// TIA Portal V21 export
// export: Created 2026-11-09T01:07:26.0249752Z, ExportSetting WithDefaults, DisplayName Totally Integrated Automation Portal, DisplayVersion V21 Update 3, DisplayName STEP 7 Professional, DisplayVersion V21 Update 3, DisplayName STEP 7 Safety, DisplayVersion V21, DisplayName Tech WebApplication, DisplayVersion V21, DisplayName WinCC Basic/Comfort/Advanced, DisplayVersion V21 Update 3, DisplayName WinCC Unified, DisplayVersion V21 Update 3
FUNCTION_BLOCK "FB_Motor"   // FB2, SCL
{ S7_Optimized_Access := 'TRUE' }
// stored: AutoNumber true, IsIECCheckEnabled false, IsRetainMemResEnabled false, MemoryReserve 100, SetENOAutomatically false, UDAEnableTagReadback false
   VAR_INPUT
      motor : "UDT_Motor";
   END_VAR
   VAR_OUTPUT
      running : Bool;
   END_VAR
BEGIN
   #running := #motor.Running;
END_FUNCTION_BLOCK
